Fanuc KAREL source: KT00760.KL

PROGRAM KT00760
%NOLOCKGROUP
VAR
  I1: INTEGER
  I2: INTEGER
  OUT: INTEGER
BEGIN
  I1 = 2
  I2 = 3
  I1 = 2
  I2 = 3
  OUT = ACOS(I1)
END KT00760
